// TIA Portal V20 export
ORGANIZATION_BLOCK "CyclicInterrupt"   // OB30, LAD, CyclicInterrupt
{ S7_Optimized_Access := 'TRUE' }
// stored: SetENOAutomatically false
   VAR_INPUT
      Initial_Call : Bool;   // Initial call of this OB
      Event_Count : Int;   // Events discarded
   END_VAR
   VAR_TEMP
      AKTUALNI_POZICE_FOLIE : DInt;
      AKTUALNI_POZICE_ETIKETA : DInt;
   END_VAR
   VAR_TEMP   // added for the SCL form of the ladder/FBD networks
      _w1 : Bool;
   END_VAR
BEGIN

REGION Network 1
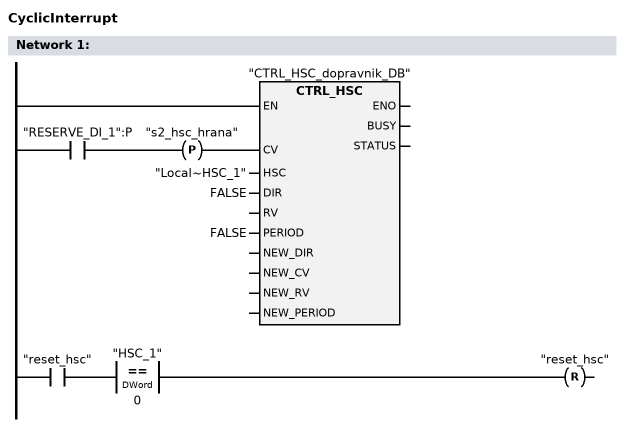
   RUNG wire#powerrail
      "CTRL_HSC_dopravnik_DB".CTRL_HSC(CV := wire#w1, HSC := "Local~HSC_1", DIR := FALSE, RV :=, PERIOD := FALSE, NEW_DIR :=, NEW_CV :=, NEW_RV :=, NEW_PERIOD :=, BUSY =>, STATUS =>)
   END_RUNG
   RUNG wire#powerrail
      Contact( "RESERVE_DI_1":P )
      P_Trig( "s2_hsc_hrana" )
   END_RUNG wire#w1
   RUNG wire#powerrail
      Contact( "reset_hsc" )
      { S7_Templates := "SrcType := DWord" } EQ_Contact(in1 := "HSC_1", in2 := 0)
      R_Coil( "reset_hsc" )
   END_RUNG
   // the same network as SCL:
   #_w1 := "RESERVE_DI_1":P AND NOT "s2_hsc_hrana";   // rising edge
   "s2_hsc_hrana" := "RESERVE_DI_1":P;
   "CTRL_HSC_dopravnik_DB"(CV := #_w1, HSC := "Local~HSC_1", DIR := FALSE, PERIOD := FALSE);   // CTRL_HSC
   IF "reset_hsc" AND ("HSC_1" = 0) THEN "reset_hsc" := FALSE; END_IF;
END_REGION

REGION Network 2 (SCL): Poloha plata od s2 [mm]
   // aktualni_poloha = HSC_1 × mm/puls (fourfold). HSC se nuluje na náběhu s2 (síť 1).
   // Konstanta 1.488 = mm na 1 puls – LIMIT brání přetečení při chodu naprázdno.
   "DB_HMI_recype".aktualni_poloha := REAL_TO_DINT(LIMIT(MN := 0.0,
                                                                                                         IN := DINT_TO_REAL(DWORD_TO_DINT("HSC_1":P)) * 4,
                                                                                                         MX := 99999.0));
END_REGION
END_ORGANIZATION_BLOCK
